// TIA Portal V20 export
Screen "Pop-up_TEC_UNIT_DIAG_LEGEND_Popup"  327x156
  ScreenItem "Background" at 0,0 size 327x156  Type=HmiRectangle
  ScreenItem "Textfeld_Legende" at 1,1 size 325x25  Type=HmiTextBox
  ScreenItem "Textfeld_3" at 10,33 size 100x20  Type=HmiTextBox
  ScreenItem "Textfeld_4" at 10,55 size 100x20  Type=HmiTextBox
  ScreenItem "Textfeld_5" at 10,103 size 100x20  Type=HmiTextBox
  ScreenItem "Textfeld_6" at 10,125 size 100x20  Type=HmiTextBox
  ScreenItem "Textfeld_11" at 115,33 size 120x20  Type=HmiTextBox
  ScreenItem "Textfeld_12" at 115,55 size 120x20  Type=HmiTextBox
  ScreenItem "Textfeld_13" at 115,103 size 120x20  Type=HmiTextBox
  ScreenItem "Textfeld_14" at 115,125 size 120x20  Type=HmiTextBox
  ScreenItem "Textfeld_15" at 10,80 size 100x20  Type=HmiTextBox
  ScreenItem "Cancel Mode" at 236,1 size 90x60  Type=HmiButton
